// Mitsubishi GX Works2 project: Tas2_Ex_3_TeachersWay   PLC: FX3G

PROGRAM MAIN
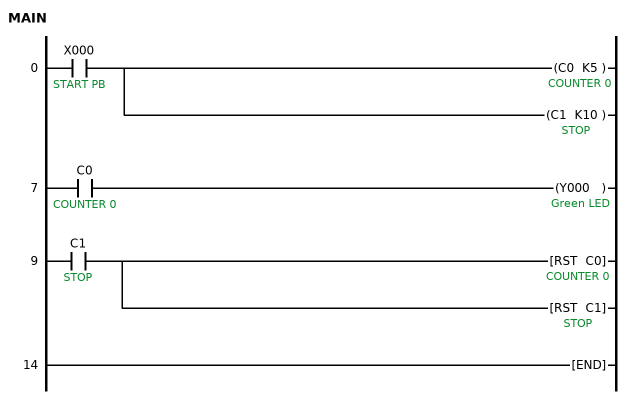
0     LD      X000  ; START PB
      OUT     C0 K5  ; COUNTER 0
      OUT     C1 K10  ; STOP
7     LD      C0  ; COUNTER 0
      OUT     Y000  ; Green LED
9     LD      C1  ; STOP
      RST     C0  ; COUNTER 0
      RST     C1  ; STOP
14    END
END_PROGRAM

// device comments not shown above
X001  ; RST
